// TIA Portal V20 export
Screen "190Passing stand"  1276x673
  ScreenItem "Line_Header_X0_Y64" at 0,64 size 1276x0  Type=HmiLine
  ScreenItem "permanentareaborderrectangle" at 0,0 size 0x0  Type=HmiRectangle
  ScreenItem "Button_Back" at 2,2 size 90x60  Type=HmiButton
  ScreenItem "Move_Legend" at 1182,2 size 90x60  Type=HmiButton
  ScreenItem "Fusszeile_Button_ManualOPMode1_2" at 100,1 size 90x60  Type=HmiButton
  ScreenItem "文本域_14" at 936,-172 size 140x40  Type=HmiTextBox
  ScreenItem "Graphic view_1" at 226,212 size 651x296  Type=HmiGraphicView
  ScreenItem "文本域_5" at -1,82 size 120x40  Type=HmiTextBox
  ScreenItem "文本域_27" at -1,126 size 120x40  Type=HmiTextBox
  ScreenItem "文本域_21" at 152,82 size 140x40  Type=HmiTextBox
  ScreenItem "Line_4" at 210,140 size 70x160  Type=HmiLine
  ScreenItem "Title_ScreenOverview_X390_Y2_1" at 384,5 size 510x57  Type=HmiTextBox
  ScreenItem "文本域_6" at 545,82 size 140x40  Type=HmiTextBox
  ScreenItem "Line_1" at 623,162 size 63x183  Type=HmiLine
  ScreenItem "文本域_7" at 879,82 size 140x40  Type=HmiTextBox
  ScreenItem "Line_2" at 808,174 size 130x206  Type=HmiLine
  ScreenItem "文本域_8" at 883,528 size 140x40  Type=HmiTextBox
  ScreenItem "面板容器_4" at 883,569 size 144x51  Type=HmiFaceplateContainer
  ScreenItem "Line_3" at 848,455 size 66x71  Type=HmiLine
  ScreenItem "文本域_9" at 72,468 size 140x40  Type=HmiTextBox
  ScreenItem "面板容器_5" at 74,509 size 144x51  Type=HmiFaceplateContainer
  ScreenItem "Line_5" at 140,336 size 121x132  Type=HmiLine
  ScreenItem "面板容器_1" at 547,125 size 144x51  Type=HmiFaceplateContainer
  ScreenItem "面板容器_8" at 154,125 size 144x51  Type=HmiFaceplateContainer
  ScreenItem "面板容器_3" at 879,125 size 144x51  Type=HmiFaceplateContainer
  ScreenItem "面板容器_2" at 1090,4 size 88x58  Type=HmiFaceplateContainer
  ScreenItem "OPMode1_Blocked" at 1164,6 size 14x14  Type=HmiGraphicView
  ScreenItem "OPMode4_Foreground_Blocked" at 1089,3 size 88x58  Type=HmiGraphicView
